(* IEC 61131-3 sources: kns-port-domestic/tools/tests/fixtures/lowering/src/POUs/PRG_Idle, 1 file *)

(* ---- PRG_Idle.decl.st ---- *)
// Назначение: пример для понижения iec-checker (tools/tests/test_assemble.py)
// Автор:      kr0nsch
// Версия:     0.1.0
// Документ:   docs/LAYOUT.md, раздел «Собранный текст build/assembled»; tools/README.md
PROGRAM PRG_Idle
VAR
    fbSlots : FB_Slots;
END_VAR
